Fanuc KAREL source: KB00057.KL

PROGRAM KB00057
%NOLOCKGROUP
VAR
  P1: INTEGER
  P2: INTEGER
BEGIN
  P1 = 1
  P2 = 1
  DAQ_UNREG(P1, P2)
END KB00057
